SUBAPPLICATION RedGreenBackground4C (* Hintergrundfarbe (TRUE -> Rot, FALSE -> Grün) für 4 Objekte (Kompakt) *)
  (* Standard: 61499-2 *)
  (* Version 1.0, 2022-11-10, franz, Meisterschulen am Ostbahnhof *)
  PACKAGE MyLib::sys;
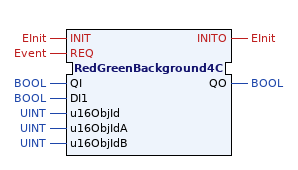
  EVENT_INPUT
    INIT : EInit; (* Initialization Request *)
    REQ; (* Normal Execution Request *)
  END_EVENT
  EVENT_OUTPUT
    INITO : EInit; (* Initialization Confirm *)
  END_EVENT
  VAR_INPUT
    QI : BOOL := TRUE; (* Quality Input - TRUE to enable service *)
    DI1 : BOOL; (* Selector *)
    u16ObjId : UINT; (* Object ID Softkey *)
    u16ObjIdA : UINT; (* Object ID AUX *)
    u16ObjIdB : UINT;
  END_VAR
  VAR_OUTPUT
    QO : BOOL; (* Quality Output - TRUE if service executed successfully *)
  END_VAR
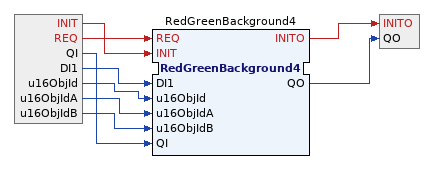
  SUBAPPS
    RedGreenBackground4 : MyLib::sys::RedGreenBackground4;
  END_SUBAPPS
  EVENT_CONNECTIONS
    REQ TO RedGreenBackground4.REQ;
    INIT TO RedGreenBackground4.INIT;
    RedGreenBackground4.INITO TO INITO;
  END_CONNECTIONS
  DATA_CONNECTIONS
    DI1 TO RedGreenBackground4.DI1;
    u16ObjId TO RedGreenBackground4.u16ObjId;
    u16ObjIdA TO RedGreenBackground4.u16ObjIdA;
    u16ObjIdB TO RedGreenBackground4.u16ObjIdB;
    QI TO RedGreenBackground4.QI;
    RedGreenBackground4.QO TO QO;
  END_CONNECTIONS
END_SUBAPPLICATION
